(* IEC 61131-3 sources: llm-plc-st-eval/data/definitivo/qwen2.5-coder_14b/B5/few_shot, 3 files *)

(* ---- ejec_1.st ---- *)
FUNCTION_BLOCK FB_Ventilador
VAR_INPUT
    quemadorOn : BOOL; (* Estado del quemador *)
END_VAR
VAR_OUTPUT
    ventilador : BOOL; (* Estado del ventilador *)
END_VAR
VAR
    tApagado : TP; (* Temporizador para el apagado *)
    estadoVentilador : BOOL; (* Estado interno del ventilador *)
END_VAR

(* Si el quemador está encendido, el ventilador también lo está *)
IF quemadorOn THEN
    estadoVentilador := TRUE;
    tApagado(IN := FALSE); (* Reiniciar el temporizador *)
ELSE
    (* Si el quemador está apagado, iniciar el temporizador *)
    tApagado(IN := TRUE, PT := T#30S);
    (* Mantener el ventilador encendido mientras el temporizador no haya expirado *)
    estadoVentilador := tApagado.Q;
END_IF;

(* Asignar el estado interno del ventilador a la salida *)
ventilador := estadoVentilador;
END_FUNCTION_BLOCK

(* ---- ejec_2.st ---- *)
FUNCTION_BLOCK FB_Ventilador
VAR_INPUT
    quemadorOn : BOOL; (* Estado del quemador *)
END_VAR
VAR_OUTPUT
    ventilador : BOOL; (* Estado del ventilador *)
END_VAR
VAR
    tApagado : TP; (* Temporizador para el apagado *)
    estadoVentilador : BOOL; (* Estado interno del ventilador *)
END_VAR

(* Si el quemador está encendido, el ventilador también lo está *)
IF quemadorOn THEN
    estadoVentilador := TRUE;
    tApagado(IN := FALSE); (* Reinicia el temporizador *)
ELSE
    (* Si el quemador está apagado, el ventilador sigue encendido durante 30 segundos *)
    tApagado(IN := TRUE, PT := T#30S);
    estadoVentilador := tApagado.Q;
END_IF;

ventilador := estadoVentilador;
END_FUNCTION_BLOCK

(* ---- ejec_3.st ---- *)
FUNCTION_BLOCK FB_Ventilador
VAR_INPUT
    quemadorOn : BOOL; (* Estado del quemador *)
END_VAR
VAR_OUTPUT
    ventilador : BOOL; (* Estado del ventilador *)
END_VAR
VAR
    tApagado : TP; (* Temporizador para el apagado *)
END_VAR

(* El ventilador funciona mientras el quemador está encendido *)
IF quemadorOn THEN
    ventilador := TRUE;
    tApagado(IN := FALSE); (* Reinicia el temporizador *)
ELSE
    (* Si el quemador está apagado, el ventilador sigue funcionando durante 30 segundos *)
    tApagado(IN := TRUE, PT := T#30S);
    ventilador := tApagado.Q;
END_IF
END_FUNCTION_BLOCK
